(* PLC project TBEN_L5_PLC11.project, CODESYS CODESYS V3.5 SP21 Patch 1 *)
(* stored: creationDateTime 2026-11-07T15:34:51.7941714, modificationDateTime 2026-11-07T15:09:07.4034196 *)

// 1 request ISDU gửi qua master
TYPE ST_IolRequest :
STRUCT
    usiPort     : USINT;                                   // 0 = master, 1..4 = port
    eService    : E_IolService := E_IolService.READ;
    uiIndex     : UINT;
    usiSubindex : USINT;                                   // 0 = cả index
    uiLen       : UINT;                                    // số byte dữ liệu ghi (READ = 0)
    abData      : ARRAY[0..GVL_IolConst.uiMAX_DATA - 1] OF BYTE;
END_STRUCT
END_TYPE
